// TIA Portal V21 export
// export: Created 2026-09-22T12:22:14.6699089Z, ExportSetting None, DisplayName Totally Integrated Automation Portal, DisplayVersion V21 Update 9, DisplayName TIA Portal Openness, DisplayVersion V21 Update 9, DisplayName TIA Portal Version Control Interface, DisplayVersion V21 Update 9, DisplayName SINAMICS Startdrive Advanced, DisplayVersion V21, DisplayName SINAMICS Startdrive G130, G150, S120, S150, SINAMICS MV, S210, DisplayVersion V21, DisplayName SINAMICS Startdrive G110M, G120, G120C, G120D, G120P, G115D, DisplayVersion V21, DisplayName STEP 7 Professional, DisplayVersion V21 Update 9, DisplayName SINUMERIK ONE STEP 7 Toolbox, DisplayVersion V21 Update 12, DisplayName SINUMERIK ONE PLC Basic Program Plus, DisplayVersion V21 Update 12, DisplayName SINUMERIK 840D sl STEP 7 Toolbox, DisplayVersion V21 Update 12, DisplayName STEP 7 Safety, DisplayVersion V21 Update 6, DisplayName WinCC Advanced, DisplayVersion V21 Update 9
FUNCTION_BLOCK "PR_ModeManageNoMode"   // FB562, LAD
TITLE = Mode Management: No mode activated during initial power on
{ S7_Optimized_Access := 'TRUE' }
AUTHOR : PARI
NAME : S11002022002
// |=============================================================================|
// BLOCK: FB601 - ModeManage_NoMode
// Item Code : S11002011002
// Owner:Precision Automation & Robotics India Ltd.
// Author: PARI
// Release Date:14-Aug-2015
// Version:0.1
// Status: Not Tested
// |=============================================================================|
// Block Description:
// This block is used Control Mode Of System.After Power On or End Of Cycle It 
// will 
// go to No Mode State if mode 
// Selection is not present
// |=============================================================================|
// 
// Dependency:
// This block uses following standard "Siemens" functions:
// SFB 4: TON : ON Delay timer
// Hence SFB4 has to be present in the CPU memory, else 
// this block call may lead to CPU going to STOP mode
// |=============================================================================|
// stored: MemoryReserve 100, SetENOAutomatically false
   VAR_INPUT
      iFirstscan : Bool;   // PLC First Scan Bit
      iControlOn : Bool;   // Machine All Safety Relay Healthy
      iAutoModeEnable : Bool;   // If conditions are OK to start automode make this bit high
      iManModeEnable : Bool;   // If conditions are OK to sart manual mode make this bit high
      iAutoMode : Bool;   // Auto Mode Input PB/SW
      iManMode : Bool;   // Man Mode Input PB/SW
      iCycleStart : Bool;   // Cycle Start Input PB
      iCycleStop : Bool;   // Cycle Stop Input PB (NC Type)
      iHomePB : Bool;   // Home Input PB
      iEndOfCycle : Bool;   // If Cycle Completed make this bit high
      iDrainCycle : Bool;   // If conditions are OK to start drain cycle make this bit high
      iDryCycle : Bool;   // If conditions are OK to start dry cycle make this bit high
      iDrainCompleted : Bool;   // If Drain Completed make this bit high
      iHomeCompleted : Bool;   // If Home Completed make this bit high
      iImmediateStop : Bool;   // To abort autocycle or to select manual while running in auto make this bit 1
      iCycleStartDelay : Time;   // Cycle Start PB Press Delay Eg. If 2Sec T#2S
      iBypassHomeOption : Bool;   // Make sure that autocycle can initiate without home condition = 1
   END_VAR
   VAR_OUTPUT
      qManModeActive : Bool;   // Man Mode Active
      qWaitForCStart : Bool;   // Waiting For Cycle Start
      qAutoRunningActive : Bool;   // AutoRunning Active
      qHomeRunningActive : Bool;   // Home Running Active
      qDrainActive : Bool;   // Drain Active
      qCycleStopActive : Bool;   // Cycle Stop Active
      qDryCycleActive : Bool;   // Dry Cycle Active
      qModuleReset : Bool;   // 1 If No Mode Selected
      qMsgCStartandNoHome : Bool;   // Cycle Start PB Pressed but MC Not at Home
      qMsgManModeinAutoRunning : Bool;   // Manual Mode selected during Auto Running
   END_VAR
   VAR
      sPowerOnReset : Bool;   // Power ON reset Bit during initial power ON
      sControlOnPulse : Bool;   // Control ON pulse
      sControlOnEdge : Bool;   // Control ON Input Positive Edge
      sManModeActivePulse : Bool;   // Man Mode Active Positive Edge Pulse
      sCycleStartDelay : Time;   // Cycle Start Delay
      CycleStartOnDelayTimer { S7_SetPoint := 'True'} : TON_TIME;   // ON Delay Timer SFB4
      sAutoRunningActive : Bool;   // Auto Running Active
      sManModeActive : Bool;   // Man Mode Active
      sHomeRunningActive : Bool;   // Home Running Active
      sWaitForCStart : Bool;   // Waiting For Cycle Start
      sDrainActive : Bool;   // Drain Active
      sDryCycleActive : Bool;   // Dry Cycle Active
      sCycleStopActive : Bool;   // Cycle Stop Active
      sModuleReset : Bool;   // Module Reset
      sMsgCStartandNoHome : Bool;   // Cycle Start PB Pressed but MC Not at Home
      sMsgManModeinAutoRunning : Bool;   // Manual Mode selected during Auto Running
   END_VAR
   VAR_TEMP   // added for the SCL form of the ladder/FBD networks
      _w1 : Bool;
      _w2 : Bool;
   END_VAR
BEGIN

REGION Network 1: Header
   // ==============================================================================
   //  Company: Precision Automation & Robotics India Ltd. 
   // ------------------------------------------------------------------------------
   //  Item Code: S11002022002
   //  Author/Created by: PARI
   //  Reviewed/Checked by: Atul P
   //  First Release on: 14-Aug-2015
   //  Latest update on: 14-Aug-2015
   // ------------------------------------------------------------------------------
   //  Tested with: CPU firmware, model or simulator testing
   //  Engineering/Editor: TIA Portal V15.1
   // ------------------------------------------------------------------------------
   //  Restrictions: No
   //  Dependencies/Requirements:
   // ------------------------------------------------------------------------------
   //  Change Log:
   //  Ver.	Date		Changed by		Details of changes
   //  1.0       14-Aug-2015                           A.D	                                     First release version
   // ------------------------------------------------------------------------------
   // Functionality:
   // This block is used Control Mode Of System.After Power On or End Of Cycle It 
   // will go to No Mode State if mode 
   // Selection is not present
   // 
   //  Inputs
   // iFirstscan	Bool
   // iContolOn	Bool
   // iAutoModeEnable	Bool
   // iManModeEnable	Bool
   // iAutoMode	Bool
   // iManMode	Bool
   // iCycleStart	Bool
   // iCycleStop	Bool
   // iHomePB	Bool
   // iEndOfCycle	Bool
   // iDrainCycle	Bool
   // iDryCycle	Bool
   // iDrainCompleted	Bool
   // iHomeCompleted	Bool
   // iImmediateStop	Bool
   // iCycleStartDelay	Time
   // iBypassHomeOption	Bool
   // 
   // 
   //  Outputs
   // qManModeActive	Bool
   // qWaitForCStart	Bool
   // qAutoRunningActive	Bool
   // qHomeRunningActive	Bool
   // qDrainActive	Bool
   // qCycleStopActive	Bool
   // qDryCycleActive	Bool
   // qModuleReset	Bool
   // 
   // 
   // In-outs
   // Nill
   // 
   // ------------------------------------------------------------------------------
   // Errors reported:
   // Nill
   // 
   // Messages:
   // qMsgCStartandNoHome	Bool
   // qMsgManModeinAutoRunning	Bool
   // 
   // ==============================================================================
END_REGION

REGION Network 2: Cycle Start delay validation
   // Cycle Start delay validation
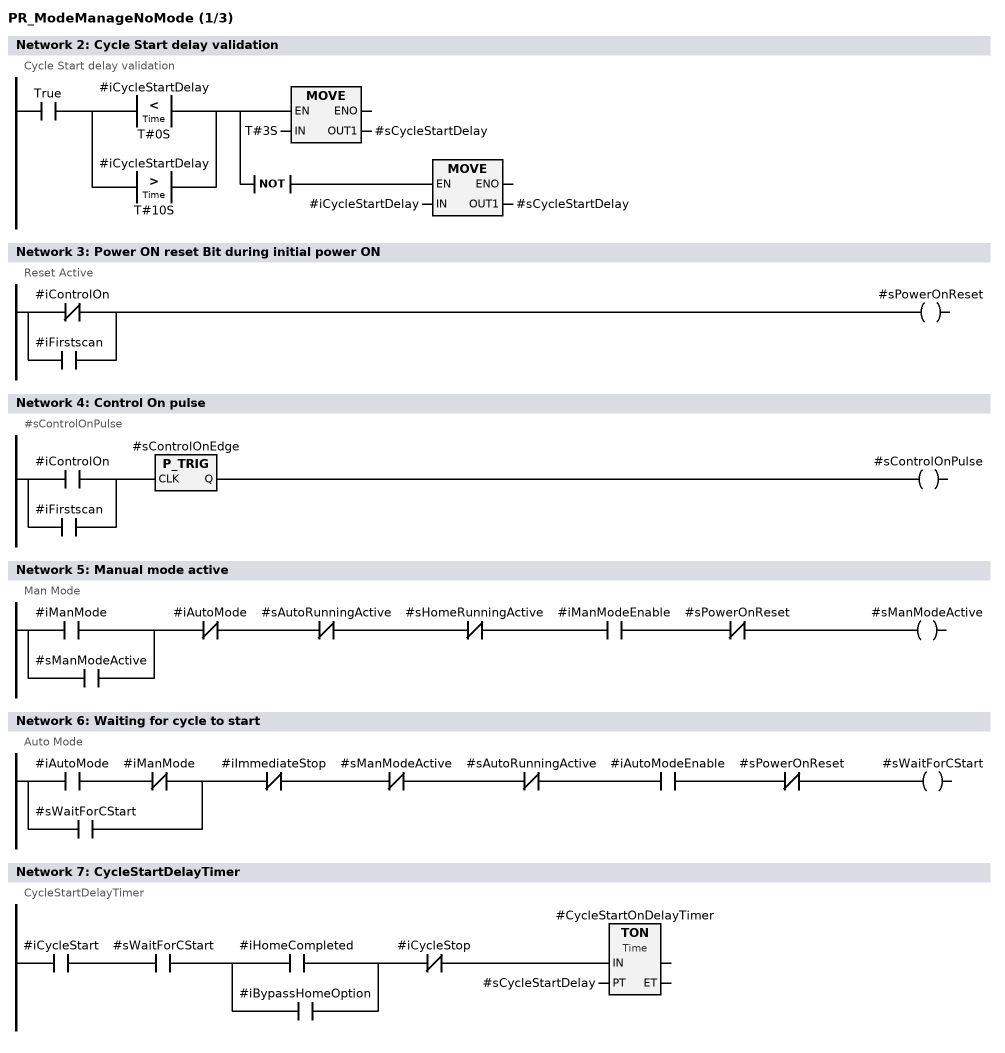
   RUNG wire#powerrail
      Contact( True )
      wire#w1
      { S7_Templates := "SrcType := Time" } LT_Contact(in1 := #iCycleStartDelay, in2 := T#0S)
      wire#w2
      Move(in := T#3S, out1 => #sCycleStartDelay)
   END_RUNG
   RUNG wire#w1
      { S7_Templates := "SrcType := Time" } GT_Contact(in1 := #iCycleStartDelay, in2 := T#10S)
   END_RUNG wire#w2
   RUNG wire#w2
      Not()
      Move(in := #iCycleStartDelay, out1 => #sCycleStartDelay)
   END_RUNG
   // the same network as SCL:
   #_w1 := True AND ((#iCycleStartDelay < T#0S) OR (#iCycleStartDelay > T#10S));
   IF #_w1 THEN #sCycleStartDelay := T#3S; END_IF;
   IF NOT #_w1 THEN #sCycleStartDelay := #iCycleStartDelay; END_IF;
END_REGION

REGION Network 3: Power ON reset Bit during initial power ON
   // Reset Active
   RUNG wire#powerrail
      I_Contact( #iControlOn )
      wire#w1
      Coil( #sPowerOnReset )
   END_RUNG
   RUNG wire#powerrail
      Contact( #iFirstscan )
   END_RUNG wire#w1
   // the same network as SCL:
   #sPowerOnReset := NOT #iControlOn OR #iFirstscan;
END_REGION

REGION Network 4: Control On pulse
   // #sControlOnPulse
   RUNG wire#powerrail
      Contact( #iControlOn )
      wire#w1
      P_Trig( #sControlOnEdge )
      Coil( #sControlOnPulse )
   END_RUNG
   RUNG wire#powerrail
      Contact( #iFirstscan )
   END_RUNG wire#w1
   // the same network as SCL:
   #_w1 := #iControlOn OR #iFirstscan;
   #_w2 := #_w1 AND NOT #sControlOnEdge;   // rising edge
   #sControlOnEdge := #_w1;
   #sControlOnPulse := #_w2;
END_REGION

REGION Network 5: Manual mode active
   // Man Mode
   RUNG wire#powerrail
      Contact( #iManMode )
      wire#w1
      I_Contact( #iAutoMode )
      I_Contact( #sAutoRunningActive )
      I_Contact( #sHomeRunningActive )
      Contact( #iManModeEnable )
      I_Contact( #sPowerOnReset )
      Coil( #sManModeActive )
   END_RUNG
   RUNG wire#powerrail
      Contact( #sManModeActive )
   END_RUNG wire#w1
   // the same network as SCL:
   #sManModeActive := (#iManMode OR #sManModeActive) AND NOT #iAutoMode AND NOT #sAutoRunningActive AND NOT #sHomeRunningActive AND #iManModeEnable AND NOT #sPowerOnReset;
END_REGION

REGION Network 6: Waiting for cycle to start
   // Auto Mode
   RUNG wire#powerrail
      Contact( #iAutoMode )
      I_Contact( #iManMode )
      wire#w1
      I_Contact( #iImmediateStop )
      I_Contact( #sManModeActive )
      I_Contact( #sAutoRunningActive )
      Contact( #iAutoModeEnable )
      I_Contact( #sPowerOnReset )
      Coil( #sWaitForCStart )
   END_RUNG
   RUNG wire#powerrail
      Contact( #sWaitForCStart )
   END_RUNG wire#w1
   // the same network as SCL:
   #sWaitForCStart := ((#iAutoMode AND NOT #iManMode) OR #sWaitForCStart) AND NOT #iImmediateStop AND NOT #sManModeActive AND NOT #sAutoRunningActive AND #iAutoModeEnable AND NOT #sPowerOnReset;
END_REGION

REGION Network 7: CycleStartDelayTimer
   // CycleStartDelayTimer
   RUNG wire#powerrail
      Contact( #iCycleStart )
      Contact( #sWaitForCStart )
      wire#w1
      Contact( #iHomeCompleted )
      wire#w2
      I_Contact( #iCycleStop )
      { S7_Templates := "time_type := Time" } #CycleStartOnDelayTimer.TON(pt := #sCycleStartDelay, et =>)
   END_RUNG
   RUNG wire#w1
      Contact( #iBypassHomeOption )
   END_RUNG wire#w2
   // the same network as SCL:
   #CycleStartOnDelayTimer(IN := #iCycleStart AND #sWaitForCStart AND (#iHomeCompleted OR #iBypassHomeOption) AND NOT #iCycleStop,   // TON
                           PT := #sCycleStartDelay);
END_REGION

REGION Network 8: Drain,Dry,Cycle Stop Active
   // Drain,Dry,Cycle Stop Active
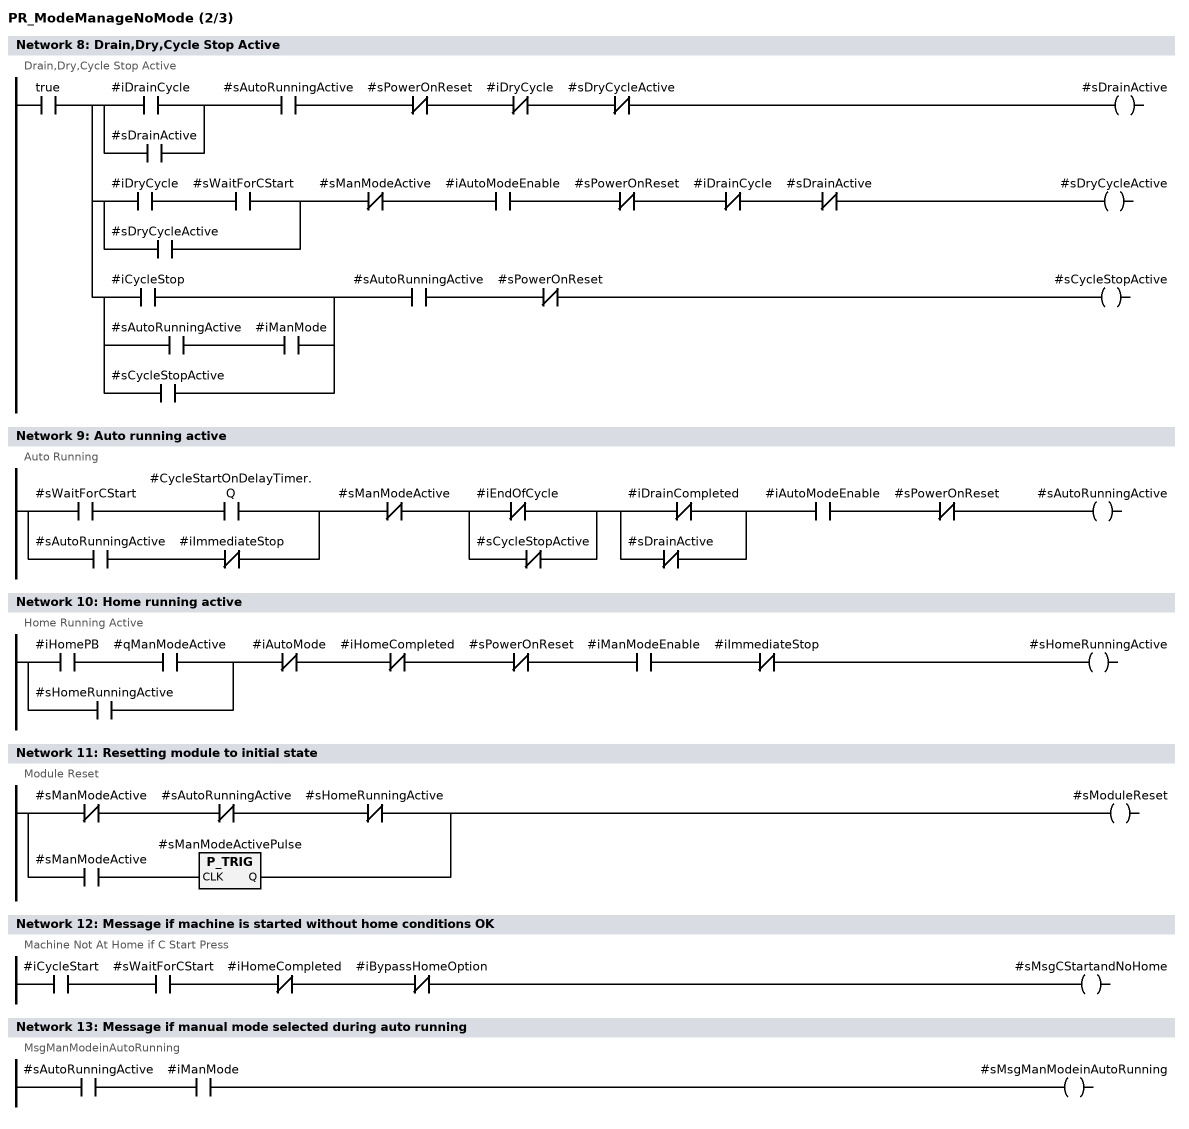
   RUNG wire#powerrail
      Contact( true )
      wire#w1
      Contact( #iDrainCycle )
      wire#w2
      Contact( #sAutoRunningActive )
      I_Contact( #sPowerOnReset )
      I_Contact( #iDryCycle )
      I_Contact( #sDryCycleActive )
      Coil( #sDrainActive )
   END_RUNG
   RUNG wire#w1
      Contact( #sDrainActive )
   END_RUNG wire#w2
   RUNG wire#w1
      Contact( #iDryCycle )
      Contact( #sWaitForCStart )
      wire#w3
      I_Contact( #sManModeActive )
      Contact( #iAutoModeEnable )
      I_Contact( #sPowerOnReset )
      I_Contact( #iDrainCycle )
      I_Contact( #sDrainActive )
      Coil( #sDryCycleActive )
   END_RUNG
   RUNG wire#w1
      Contact( #sDryCycleActive )
   END_RUNG wire#w3
   RUNG wire#w1
      Contact( #iCycleStop )
      wire#w4
      Contact( #sAutoRunningActive )
      I_Contact( #sPowerOnReset )
      Coil( #sCycleStopActive )
   END_RUNG
   RUNG wire#w1
      Contact( #sAutoRunningActive )
      Contact( #iManMode )
   END_RUNG wire#w4
   RUNG wire#w1
      Contact( #sCycleStopActive )
   END_RUNG wire#w4
   // the same network as SCL:
   #sDrainActive := true AND (#iDrainCycle OR #sDrainActive) AND #sAutoRunningActive AND NOT #sPowerOnReset AND NOT #iDryCycle AND NOT #sDryCycleActive;
   #sDryCycleActive := true AND ((#iDryCycle AND #sWaitForCStart) OR #sDryCycleActive) AND NOT #sManModeActive AND #iAutoModeEnable AND NOT #sPowerOnReset AND NOT #iDrainCycle AND NOT #sDrainActive;
   #sCycleStopActive := true AND (#iCycleStop OR (#sAutoRunningActive AND #iManMode) OR #sCycleStopActive) AND #sAutoRunningActive AND NOT #sPowerOnReset;
END_REGION

REGION Network 9: Auto running active
   // Auto Running
   RUNG wire#powerrail
      Contact( #sWaitForCStart )
      Contact( #CycleStartOnDelayTimer.Q )
      wire#w1
      I_Contact( #sManModeActive )
      wire#w2
      I_Contact( #iEndOfCycle )
      wire#w3
      I_Contact( #iDrainCompleted )
      wire#w4
      Contact( #iAutoModeEnable )
      I_Contact( #sPowerOnReset )
      Coil( #sAutoRunningActive )
   END_RUNG
   RUNG wire#powerrail
      Contact( #sAutoRunningActive )
      I_Contact( #iImmediateStop )
   END_RUNG wire#w1
   RUNG wire#w2
      I_Contact( #sCycleStopActive )
   END_RUNG wire#w3
   RUNG wire#w3
      I_Contact( #sDrainActive )
   END_RUNG wire#w4
   // the same network as SCL:
   #sAutoRunningActive := ((#sWaitForCStart AND #CycleStartOnDelayTimer.Q) OR (#sAutoRunningActive AND NOT #iImmediateStop)) AND NOT #sManModeActive AND (NOT #iEndOfCycle OR NOT #sCycleStopActive) AND (NOT #iDrainCompleted OR NOT #sDrainActive) AND #iAutoModeEnable AND NOT #sPowerOnReset;
END_REGION

REGION Network 10: Home running active
   // Home Running Active
   RUNG wire#powerrail
      Contact( #iHomePB )
      Contact( #qManModeActive )
      wire#w1
      I_Contact( #iAutoMode )
      I_Contact( #iHomeCompleted )
      I_Contact( #sPowerOnReset )
      Contact( #iManModeEnable )
      I_Contact( #iImmediateStop )
      Coil( #sHomeRunningActive )
   END_RUNG
   RUNG wire#powerrail
      Contact( #sHomeRunningActive )
   END_RUNG wire#w1
   // the same network as SCL:
   #sHomeRunningActive := ((#iHomePB AND #qManModeActive) OR #sHomeRunningActive) AND NOT #iAutoMode AND NOT #iHomeCompleted AND NOT #sPowerOnReset AND #iManModeEnable AND NOT #iImmediateStop;
END_REGION

REGION Network 11: Resetting module to initial state
   // Module Reset
   RUNG wire#powerrail
      I_Contact( #sManModeActive )
      I_Contact( #sAutoRunningActive )
      I_Contact( #sHomeRunningActive )
      wire#w1
      Coil( #sModuleReset )
   END_RUNG
   RUNG wire#powerrail
      Contact( #sManModeActive )
      P_Trig( #sManModeActivePulse )
   END_RUNG wire#w1
   // the same network as SCL:
   #_w1 := #sManModeActive AND NOT #sManModeActivePulse;   // rising edge
   #sManModeActivePulse := #sManModeActive;
   #sModuleReset := (NOT #sManModeActive AND NOT #sAutoRunningActive AND NOT #sHomeRunningActive) OR #_w1;
END_REGION

REGION Network 12: Message if machine is started without home conditions OK
   // Machine Not At Home if C Start Press
   RUNG wire#powerrail
      Contact( #iCycleStart )
      Contact( #sWaitForCStart )
      I_Contact( #iHomeCompleted )
      I_Contact( #iBypassHomeOption )
      Coil( #sMsgCStartandNoHome )
   END_RUNG
   // the same network as SCL:
   #sMsgCStartandNoHome := #iCycleStart AND #sWaitForCStart AND NOT #iHomeCompleted AND NOT #iBypassHomeOption;
END_REGION

REGION Network 13: Message if manual mode selected during auto running
   // MsgManModeinAutoRunning
   RUNG wire#powerrail
      Contact( #sAutoRunningActive )
      Contact( #iManMode )
      Coil( #sMsgManModeinAutoRunning )
   END_RUNG
   // the same network as SCL:
   #sMsgManModeinAutoRunning := #sAutoRunningActive AND #iManMode;
END_REGION

REGION Network 14: Outputs
   // Outputs
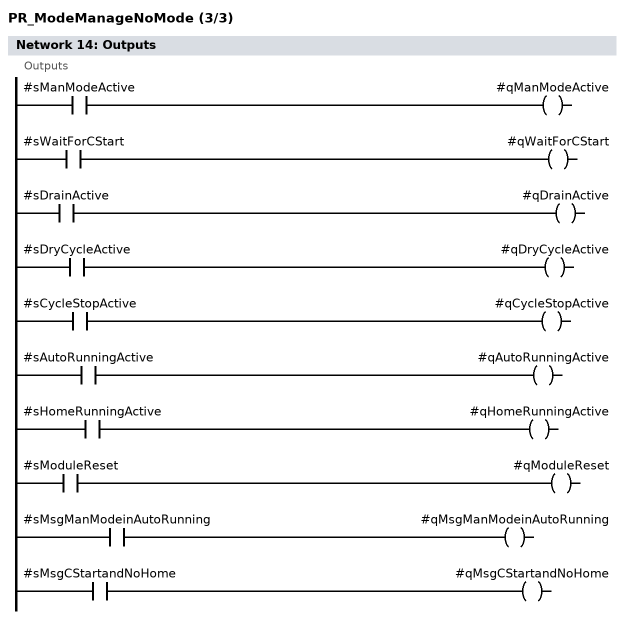
   RUNG wire#powerrail
      Contact( #sManModeActive )
      Coil( #qManModeActive )
   END_RUNG
   RUNG wire#powerrail
      Contact( #sWaitForCStart )
      Coil( #qWaitForCStart )
   END_RUNG
   RUNG wire#powerrail
      Contact( #sDrainActive )
      Coil( #qDrainActive )
   END_RUNG
   RUNG wire#powerrail
      Contact( #sDryCycleActive )
      Coil( #qDryCycleActive )
   END_RUNG
   RUNG wire#powerrail
      Contact( #sCycleStopActive )
      Coil( #qCycleStopActive )
   END_RUNG
   RUNG wire#powerrail
      Contact( #sAutoRunningActive )
      Coil( #qAutoRunningActive )
   END_RUNG
   RUNG wire#powerrail
      Contact( #sHomeRunningActive )
      Coil( #qHomeRunningActive )
   END_RUNG
   RUNG wire#powerrail
      Contact( #sModuleReset )
      Coil( #qModuleReset )
   END_RUNG
   RUNG wire#powerrail
      Contact( #sMsgManModeinAutoRunning )
      Coil( #qMsgManModeinAutoRunning )
   END_RUNG
   RUNG wire#powerrail
      Contact( #sMsgCStartandNoHome )
      Coil( #qMsgCStartandNoHome )
   END_RUNG
   // the same network as SCL:
   #qManModeActive := #sManModeActive;
   #qWaitForCStart := #sWaitForCStart;
   #qDrainActive := #sDrainActive;
   #qDryCycleActive := #sDryCycleActive;
   #qCycleStopActive := #sCycleStopActive;
   #qAutoRunningActive := #sAutoRunningActive;
   #qHomeRunningActive := #sHomeRunningActive;
   #qModuleReset := #sModuleReset;
   #qMsgManModeinAutoRunning := #sMsgManModeinAutoRunning;
   #qMsgCStartandNoHome := #sMsgCStartandNoHome;
END_REGION
END_FUNCTION_BLOCK
